// TIA Portal V20 export
// export: Created 2026-11-12T11:17:33.9952123Z, ExportSetting WithDefaults, DisplayName Totally Integrated Automation Portal, DisplayVersion V20, DisplayName TIA Portal Openness, DisplayVersion V20, DisplayName TIA Portal Teamcenter Gateway, DisplayVersion V20, DisplayName TIA Portal Version Control Interface, DisplayVersion V20, DisplayName STEP 7 Professional, DisplayVersion V20, DisplayName STEP 7 CFC, DisplayVersion V20, DisplayName STEP 7 Safety, DisplayVersion V20, DisplayName WinCC Basic/Comfort/Advanced, DisplayVersion V20, DisplayName SIMATIC Visualization Architect, DisplayVersion V20, DisplayName WinCC Professional, DisplayVersion V20, DisplayName SIMATIC Visualization Architect, DisplayVersion V20, DisplayName WinCC Unified, DisplayVersion V20, DisplayName SIMATIC Visualization Architect, DisplayVersion V20
TYPE "UDT_Salidas_RFID"
// stored: IsFailsafeCompliant false
   STRUCT
      Tag_escribir : Bool;   // Escribir en tag
      Tag_leer : Bool;   // Leer de tag
      Tag_reservado_2 : Bool;   // xBit2
      Tag_reservado_3 : Bool;   // xBit3
      Tag_antena_apagar : Bool;   // Apagar antena
      Tag_reservado_5 : Bool;   // xBit5
      Tag_reservado_6 : Bool;   // xBit6
      Tag_reservado_7 : Bool;   // xBit7
      Reservado_AB5 : Byte;   // byReserved
      Tag_direccion_leer_escribir : Word;   // Direccion de R/W
      Tag_datos_a_escribir : Array[0..27] of Byte;   // Datos a escribir
   END_STRUCT;
END_TYPE
